(* IEC 61131-3 sources: SortJet_MasterSPS_Aufbau.fbsproj/10_Schnittstellen, 8 files *)

(* ---- Auftragswarteschlange_Fremdanlage_FB.fb.st ---- *)
(* METADATA
{
	"v3Meta": {
		"objectGuid": "565d8e9e-6f44-455e-86f5-d16ff6a06f95"
	}
}
*)
FUNCTION_BLOCK Auftragswarteschlange_Fremdanlage_FB
VAR_INPUT

  bpAktivieren     : BOOL := TRUE;
  bpWertAuslesen   : BOOL; // READ
  bpWerteSchreiben : BOOL; // WRITE
  bpReset          : BOOL; // RST

  // WORD
  ppEingabeWert : Schnittstelle_Auftragsdaten_ST;

END_VAR
VAR_OUTPUT
  // BOOLEAN
  bpWarteschlangeLeer  : BOOL := TRUE;
  bpWarteschlangeVoll  : BOOL;

  // STRUCT
  ppAusgabeWert  : Schnittstelle_Auftragsdaten_ST;

END_VAR
VAR

  // STRUCT
  awlWarteSchlange : ARRAY[0..cINDEX] OF Schnittstelle_Auftragsdaten_ST;

  // INT
  ilAktuellePosition  : INT; // pr
  ilLetztePosition    : INT; // pw

END_VAR

VAR CONSTANT
  cINDEX : INT := 5;    // WICHTIG: Aenderungen an diesem Wert aendert die Anzahl der Elemente in der Warteschlange [FIFO]
END_VAR
IF ( bpReset ) THEN
  ilLetztePosition := ilAktuellePosition := 0 ;
  bpWarteschlangeVoll := FALSE;
  bpWarteschlangeLeer := TRUE;

  bpReset := FALSE;

ELSIF ( bpAktivieren ) THEN

  IF (  NOT bpWarteschlangeLeer
       AND bpWertAuslesen )
  THEN
    ppAusgabeWert := awlWarteSchlange[ilAktuellePosition];
    ilAktuellePosition  := INCI(ilAktuellePosition,cINDEX);
    bpWarteschlangeLeer := ilAktuellePosition = ilLetztePosition;
    bpWarteschlangeVoll := FALSE;
    bpWertAuslesen      := FALSE;
  END_IF;

  IF (  NOT bpWarteschlangeVoll
       AND bpWerteSchreiben )
  THEN
    awlWarteSchlange[ilLetztePosition] := ppEingabeWert;
    ilLetztePosition    := INCI(ilLetztePosition,cINDEX);
    bpWarteschlangeVoll := ilLetztePosition = ilAktuellePosition;
    bpWarteschlangeLeer := FALSE;
    bpWerteSchreiben    := FALSE;
  END_IF;

END_IF;
END_FUNCTION_BLOCK

(* ---- Schnittstelle_Auslauf_ISO_FB.fb.st ---- *)
(* METADATA
{
	"v3Meta": {
		"objectGuid": "159241df-4e26-44a3-b242-7f4886765264"
	}
}
*)
FUNCTION_BLOCK Schnittstelle_Auslauf_ISO_FB EXTENDS Basic_Schnittstelle_FB_V01_00_00

VAR_INPUT
END_VAR
VAR_OUTPUT
END_VAR
VAR

  // STEPS
  steplStartIsolinie       : Steps_TE;

  // TRIGGER
  rtlAutomatik             : R_TRIG;
  rtlGlasAbruf             : R_TRIG;
  ftlGlasAbruf             : F_TRIG;

END_VAR

VAR_INPUT

  // HARDWARE EINGAENGE
  in_bGlasAbruf                 AT%I* : BOOL; // Signal von ISO-Linie
  in_bTransportRueckwaerts      AT%I* : BOOL; // Signal von ISO-Linie

  // ANALOGWERT
  in_wAnalogwertISOLinie        AT%I* : WORD; // Geschwindigkeit von der ISO-Linie

END_VAR

//-------------------------------------------------------------------------------------------------
// MASTER AUFRUFEN
//-------------------------------------------------------------------------------------------------
SUPER^(BasisStationsParameter := BasisStationsParameter);

//-------------------------------------------------------------------------------------------------
// BAUSTEIN: DEAKTIVIERUNG
//-------------------------------------------------------------------------------------------------
(* Hinweis:
   - Schnittstelle deaktiviert (MK bDeaktivieren): Baustein verlassen (Ausgaenge schaltet der Basis-Baustein ab)
*)
IF ( BasisStationsParameter.stMKs.bDeaktivieren ) THEN
  RETURN;
END_IF

//-------------------------------------------------------------------------------------------------
// BAUSTEIN: AKTIONEN
//-------------------------------------------------------------------------------------------------
CASE BasisStationsParameter.stMKs.stFremdanlage.eTypSchnittstelle OF

  //eGlaston:
  //  Glaston_Schnittstelle();

  eLISEC:
    Lisec_Schnittstelle();

  eFOREL:
    Forel_Schnittstelle();

  eHEGLA_SJ:
    Hegla_SJ_Schnittstelle();

END_CASE

// Meldung: Glas bereit, aber kein Abruf durch die Fremdanlage
Meldungen();

// Glaettung der Geschwindigkeit zur Sortierung
M_GeschwindigkeitGlaetten( rpMindestGeschwindigkeitsAenderung   := BasisStationsParameter.stMKs.stFremdanlage.rMindestGeschwindigkeitsAenderung,
                           tpMindestZeitZwischenGeschwAenderung := BasisStationsParameter.stMKs.stFremdanlage.tMindestZeitZwischenGeschwAenderung );

IF BasisStationsParameter.stMKs.stFremdanlage.bStationStatusZuGlasAbruf THEN
  Status_ISO_Linie();
END_IF

IF BasisStationsParameter.stMKs.stFremdanlage.bSignaleLoggen THEN
  Signal_Logger();
END_IF
END_FUNCTION_BLOCK

(* ---- Schnittstelle_Auslauf_Schneidanlage.fb.st ---- *)
(* METADATA
{
	"v3Meta": {
		"objectGuid": "5c116975-7ea8-4794-b20d-23cbba1de39f"
	}
}
*)
FUNCTION_BLOCK Schnittstelle_Auslauf_Schneidanlage EXTENDS Basic_Schnittstelle_FB_V01_00_00

VAR_INPUT
END_VAR

VAR_OUTPUT

  // Bool
  bpAnforderungSK : BOOL;
  bpGlasAbruf     : BOOL;

END_VAR

VAR

END_VAR

VAR_INPUT

  // HARDWARE EINGAENGE
  in_bGlasAbruf                 AT%I* : BOOL; // Signal von Schneidanlage
  in_bAnforderungSK             AT%I* : BOOL; // Signal von Schneidanlage

  out_bFreigabeSK               AT%Q* : BOOL; // Signal an Schneidanlage

END_VAR

//-------------------------------------------------------------------------------------------------
// MASTER AUFRUFEN
//-------------------------------------------------------------------------------------------------
SUPER^(BasisStationsParameter := BasisStationsParameter);

//-------------------------------------------------------------------------------------------------
// BAUSTEIN: DEAKTIVIERUNG
//-------------------------------------------------------------------------------------------------
(* Hinweis:
   - Schnittstelle deaktiviert (MK bDeaktivieren): Ausgaenge abschalten, Baustein verlassen
*)
IF ( BasisStationsParameter.stMKs.bDeaktivieren ) THEN
  out_bFreigabeSK := FALSE;
  bpAnforderungSK := FALSE;
  bpGlasAbruf     := FALSE;
  RETURN;
END_IF

//-------------------------------------------------------------------------------------------------
// BAUSTEIN: AKTIONEN
//-------------------------------------------------------------------------------------------------

Signalverarbeitung();
IF BasisStationsParameter.stMKs.stFremdanlage.bSignaleLoggen THEN
  Signal_Logger();
END_IF

//-------------------------------------------------------------------------------------------------
// STEUERUNG: HARDWARESCHNITTSTELLE
//-------------------------------------------------------------------------------------------------
blSenderGlasBereit := ( (*( BasisStationsParameter.bAutomatik )
                        AND*) NOT BasisStationsParameter.InGlasTransportVorgaenger[cWAND_1].bFehler )
                      AND ( BasisStationsParameter.InGlasTransportVorgaenger[cWAND_1].bBereitZumAustransport
                            OR BasisStationsParameter.bCheckMitVorgaenger[cWAND_1]
                            OR BasisStationsParameter.bCheckMitNachfolger[cWAND_1] );

bpAnforderungSK := in_bAnforderungSK OR bgVisu_Schnittstelle_Force_AnforderungSK[BasisStationsParameter.stMKs.stStationsNummern.NummerSPS];
bpGlasAbruf     := in_bGlasAbruf OR bgVisu_Schnittstelle_Force_GlasAbruf[BasisStationsParameter.stMKs.stStationsNummern.NummerSPS];

// SK-Freigabe an die Schneidanlage: nur auf Anforderung und bei Freigabe der Schnittstelle
out_bFreigabeSK := bpAnforderungSK AND BasisStationsParameter.stFreigabe.bAlles;

bgVisu_Schnittstelle_GlasAbruf[BasisStationsParameter.stMKs.stStationsNummern.NummerSPS]     := in_bGlasAbruf OR bgVisu_Schnittstelle_Force_GlasAbruf[BasisStationsParameter.stMKs.stStationsNummern.NummerSPS];
bgVisu_Schnittstelle_AnforderungSK[BasisStationsParameter.stMKs.stStationsNummern.NummerSPS] := in_bAnforderungSK OR bgVisu_Schnittstelle_Force_AnforderungSK[BasisStationsParameter.stMKs.stStationsNummern.NummerSPS];
bgVisu_Schnittstelle_FreigabeSK[BasisStationsParameter.stMKs.stStationsNummern.NummerSPS]    := out_bFreigabeSK;
END_FUNCTION_BLOCK

(* ---- Schnittstelle_Auslauflinie_Glaston_Koppler_FB.fb.st ---- *)
(* METADATA
{
	"v3Meta": {
		"objectGuid": "1b8cd41b-c6ec-4747-8cfe-b17b04789a14"
	}
}
*)
FUNCTION_BLOCK Schnittstelle_Auslauflinie_Glaston_Koppler_FB  EXTENDS Basic_Schnittstelle_FB_V01_00_00

VAR_INPUT

  // BOOL
  bpAuftragsdatenVorhanden  : BOOL;

  // STRUCT
  Auftragsdaten             : Schnittstelle_Auftragsdaten_ST;

END_VAR
VAR_OUTPUT

END_VAR
VAR

  // BOOL
  bpDatenformatASCII                      : BOOL := TRUE;
  blLiveCounterGueltig                    : BOOL;
  blFehlermeldungGenerierenKommunikation  : BOOL;
  blFehlermeldungGenerierenAuftragsdaten  : BOOL;
  bpFehlerMeldungDeaktiviert              : BOOL := FALSE;

  // BYTE
  aOutByteLadeID             : ARRAY [0..15] OF BYTE; // Visualisierung: Lade-ID byteweise

  // WORD
  wlVerbindungsVersuche      : WORD;
  wlLiveCounterSortJet       : WORD;
  wlLiveCounterFremdanlage   : WORD;
  wlTempEmpfaengerSignale    : WORD;
  wlTempSenderSignale        : WORD;
  wlOutSignale               : WORD;
  wlInSignale                : WORD;

  // DWORD
  dwlGeschwindigkeit         : DWORD;                   // Geschwindigkeit des Empfaengers [mm/s], ggf. geswappt
  adwlLadeID                 : ARRAY [0..3] OF DWORD;   // Lade-ID (= Scheiben-ID 1), ggf. geswappt

  // INT
  ilIndex                    : INT;

  // TRIGGER
  ftlGlasBereit                           : F_TRIG; // Hinweis: Glas-Sender besitzt noch einen aktiven Transport-Zustand
  ftlFremdanlageDatenVerarbeitet          : F_TRIG;
  rtlFehlermeldungGenerierenAuftragsdaten : R_TRIG;
  rtlFehlermeldungGenerierenKommunikation : R_TRIG;

  // TIMER
  tonlZeitLiveCounterNichtAequivalent     : TON;
  tonlZeitLiveCounterInkrementieren       : TON;
  tonlZeitAuftragsdatenNichtAequivalent   : TON;
  tonlManuellerModus                      : TON;
  tonlAuftragdatenVorhanden               : TON;

  // STRING
  strScheibenID  : STRING;

  // STRUCT
  stlAuftragsdatenLeer : Schnittstelle_Auftragsdaten_ST; // Leere Auftragsdaten zum Loeschen beim Reset

  // REFERENZ
  stlVorgaenger  : REFERENCE TO StationBasisParameter_ST; // SortJet- Station vor der Schnittstelle (SF/SB)

END_VAR

VAR

  // STEPS
  steplStartIsolinie                                     : Steps_TE;

  // TRIGGER
  rtlAutomatik                                           : R_TRIG;
  rtlGlasAbruf                                           : R_TRIG;
  ftlGlasAbruf                                           : F_TRIG;

  // HARDWARE EINGAENGE KOPPLER (Hegla Schnittstellenbeschreibung V4.0, Empfaenger -> Sender)
  in_wEmpfaengerLiveCounter                     AT %I*   : WORD;                  // Wort 0     LC: gespiegelter LiveCounter
  in_awEmpfaengerLadeIDGespiegelt               AT %I*   : ARRAY [1..8] OF WORD;  // Wort 1..8  ID: gespiegelte Lade-ID
  in_wEmpfaengerSignale                         AT %I*   : WORD;                  // Wort 49    Signale
  in_dwEmpfaengerGeschwindigkeit                AT %I*   : DWORD;                 // Wort 50    GE: Geschwindigkeit [mm/s]
  in_wEmpfaengerRampe                           AT %I*   : WORD;                  // Wort 52    RA [Option]: Rampe [mm/s²], nur Anzeige

  in_bEmpfaengerAuftragsdatenErhalten                    : BOOL; // 49.0 AG
  in_bEmpfaengerBereitZumEintransport                    : BOOL; // 49.1 GA
  in_bEmpfaengerNothalt                                  : BOOL; // 49.3 NA  [Option] nur Anzeige
  in_bEmpfaengerAnforderungDurchgangOeffnen              : BOOL; // 49.4 ADO [Option] nur Anzeige
  in_bEmpfaengerQuittungDurchgangOeffnen                 : BOOL; // 49.5 ADQ [Option] nur Anzeige
  in_bEmpfaengerStationFrei                              : BOOL; // 49.6 SF  [Option]
  in_bEmpfaengerStationBeladen                           : BOOL; // 49.7 SB  [Option]
  in_bEmpfaengerUebernahmeposition                       : BOOL; // 49.8 UP  [Option] nur Anzeige

  // HARDWARE AUSGAENGE KOPPLER (Hegla Schnittstellenbeschreibung V4.0, Sender -> Empfaenger)
  out_wSenderLiveCounter                     AT %Q*      : WORD;                  // Wort 0     LC: LiveCounter
  out_awSenderLadeID                         AT %Q*      : ARRAY [1..8] OF WORD;  // Wort 1..8  ID: Lade-ID (16 ASCII- Zeichen)
  out_wSenderSignale                         AT %Q*      : WORD;                  // Wort 50    Signale

  out_bSenderAuftragdatenVorhanden                       : BOOL; // 50.0 AV
  out_bSenderAuftragdatenPlausibel                       : BOOL; // 50.1 AP
  out_bSenderManuelleBeladung                            : BOOL; // 50.2 HB [Option] SortJet sendet immer mit Lade-ID
  out_bSensorAuslauf                                     : BOOL; // 50.6 SA [Option]
  out_bSenderStationFrei                                 : BOOL; // 50.7 SF [Option] Vorgaengerstation frei
  out_bSenderStationBeladen                              : BOOL; // 50.8 SB [Option] Vorgaengerstation belegt
  out_bSenderForm                                        : BOOL; // 50.9 FG [Option] Scheibe ist ein Modell

END_VAR
VAR CONSTANT

  // WORD
  cVERBINDUNGSVERSUCHE_BIS_FEHLER  : WORD := 5;         // WICHTIG: Aenderung an diesem Wert veraendert das Verhalten ab wieviel Kommunikations-Versuchen wann ein Fehler ausgegeben wird

  // INT
  cWERTEBREICH_INT                 : INT  := 32767; // WICHTIG: Aenderung an diesem Wert aendert den Wertebereich eines INTs [positiver Wertebereich]
  cWERTEBREICH_WORD                : WORD := 32767; // WICHTIG: Aenderung an diesem Wert aendert den Wertebereich eines INTs [positiver Wertebereich]

  // TIME
  cZEIT_AUFTRAGSDATEN_GUELTIG                : TIME :=T#5s;         // WICHTIG: Aenderung an diesem Wert aendert die Zeit ab wann ein Fehlergeneriert wird [s]
  cZEIT_GESPIEGELTE_AUFTRAGSDATEN_UNGUELTIG  : TIME :=T#5s;         // WICHTIG: Aenderung an diesem Wert aendert die Zeit ab wann ein Fehlergeneriert wird [s]
  cZEIT_MANUELLER_MODUS_SIGNAL               : TIME :=T#10s;
  cZEIT_LIVECOUNTER_INKREMENTIEREN           : TIME :=T#250ms;
  cZEIT_LIVECOUNTER_NICHT_GUELTIG            : TIME :=T#1500ms;

END_VAR
//-------------------------------------------------------------------------------------------------
// MASTER AUFRUFEN
//-------------------------------------------------------------------------------------------------
SUPER^(BasisStationsParameter := BasisStationsParameter);

//-------------------------------------------------------------------------------------------------
// BAUSTEIN: INITIALISIERUNG
//-------------------------------------------------------------------------------------------------
IF ( blErsterZyklus  ) THEN
  blErsterZyklus := FALSE;

  bpAuftragsdatenVorhanden      := FALSE;
  AuftragsSpeicher.bpAktivieren := TRUE;

END_IF

//-------------------------------------------------------------------------------------------------
// BAUSTEIN: DEAKTIVIERUNG
//-------------------------------------------------------------------------------------------------
(* Hinweis:
   - Schnittstelle deaktiviert (MK bDeaktivieren): Signalwort zum Empfaenger nullen, Baustein verlassen
     (der LiveCounter bleibt stehen -> Empfaenger erkennt die fehlende Kommunikation)
*)
IF ( BasisStationsParameter.stMKs.bDeaktivieren ) THEN
  out_wSenderSignale := 0;
  RETURN;
END_IF

//-------------------------------------------------------------------------------------------------
// TIMER
//-------------------------------------------------------------------------------------------------
(* Hinweis:
   - Zeitlicheueberwachung der Kommunikation
*)
tonlZeitLiveCounterNichtAequivalent( IN := NOT blLiveCounterGueltig,
                                     PT := cZEIT_LIVECOUNTER_NICHT_GUELTIG );

//-------------------------------------------------------------------------------------------------
// AKTIONEN
//-------------------------------------------------------------------------------------------------
LiveCounter();
Meldungen();
AuftragsdatenVerwaltung();
Auswertung();
Signalverarbeitung();
M_GeschwindigkeitGlaetten( rpMindestGeschwindigkeitsAenderung   := BasisStationsParameter.stMKs.stFremdanlage.rMindestGeschwindigkeitsAenderung,
                           tpMindestZeitZwischenGeschwAenderung := BasisStationsParameter.stMKs.stFremdanlage.tMindestZeitZwischenGeschwAenderung );
Status_ISO_Linie();

IF BasisStationsParameter.stMKs.stFremdanlage.bSignaleLoggen THEN
  Signal_Logger();
END_IF

//-------------------------------------------------------------------------------------------------
// RESET
//-------------------------------------------------------------------------------------------------
// Fehlverhalten:
//   - Anstehenden Fehler zuruecksetzen
IF ( BasisStationsParameter.bReset ) THEN

  out_bSenderAuftragdatenPlausibel := FALSE;
  out_bSenderAuftragdatenVorhanden := FALSE;

  bpAuftragsdatenVorhanden               := FALSE;
  blFehlermeldungGenerierenKommunikation := FALSE;
  blFehlermeldungGenerierenAuftragsdaten := FALSE;

  BasisStationsParameter.bReset := FALSE;

  // Auftragsdaten komplett loeschen
  Auftragsdaten := stlAuftragsdatenLeer;

END_IF

//-------------------------------------------------------------------------------------------------
// Aufrufe
//-------------------------------------------------------------------------------------------------
Horn( bpAktiv := bgHornAktivieren );
END_FUNCTION_BLOCK

(* ---- Schnittstelle_Einlauf_HeglaBrechanlage_FB.fb.st ---- *)
(* METADATA
{
	"v3Meta": {
		"objectGuid": "887b7e5f-63a1-4543-befe-d3acd4ce4d49"
	}
}
*)
{attribute 'excludefrombuild'}
FUNCTION_BLOCK Schnittstelle_Einlauf_HeglaBrechanlage_FB
(*
//=================================================================================================
// !!! TODO !!! TODO !!! TODO !!! TODO !!! TODO !!! TODO !!! TODO !!! TODO !!! TODO !!! TODO !!!
//=================================================================================================
// - Dieser Baustein erbt NICHT von Basic_Schnittstelle_FB_V01_00_00.
// - Er ist nicht instanziiert und nicht im Build (excludefrombuild).
// - Vor der Verwendung auf die Basis-Schnittstelle umstellen:
//     EXTENDS, SUPER^, Reset und Meldungen der Basis nutzen, danach testen.
//=================================================================================================
*)
VAR_INPUT

  // BOOL
  bpStarteReset                 : BOOL;
  bpAnforderungSK               : BOOL;

  // STRUCT
  InGlasTransportNachfolger     : Interface_GlasTransport;
  stStationsNummern             : Station_ST;

  // POINTER
  ppParameterBaustein : REFERENCE TO Parameter_Schnittstelle;

END_VAR
VAR_OUTPUT

  // STRUCT
  OutGlasTransport : Interface_GlasTransport; // STRUKTUR: Informationen ueber den Aus- Ein- Transport WAND 1

END_VAR
VAR

  // BOOL
  blErsterZyklus          : BOOL := TRUE;

  // TIMER
  tonlMeldungGenerierenGLassenderNichtBereit : TON;// EINSCHALTVERZOEGERUNG

END_VAR
VAR

  // HARDWARE EINGAENGE
  in_bGlasBereit                AT %I* : BOOL; // Glas auf Brechanlage bereit zum Austransport
  in_bFreigabeSK                AT %I* : BOOL; // Freigabe zum SK 2 öffnen
  in_bAnlageEingeschaltet       AT %I* : BOOL; // Signal zum Zustand der Brechanlage, ob Eingeschaltet oder nicht
  in_bSensorAuslauf             AT %I* : BOOL; // Auslaufsensor (letzter Sensor vor Übergabe) der Brechanlage
  in_bBypassMode                AT %I* : BOOL; // ByPass an Brechanlage aktiv: Übergroße Scheiben für die Brechanlage müssen ohne Analogwert gefahren werden ; Festgesetzte Geschw. 20m/min zwischen Brechanlage und SortJet

  // HARDWARE AUSGAENGE
  out_bGlasAbruf                AT %Q* : BOOL; // Glas Abruf zur Brechanlage, sofern Glas Bereit ist
  out_bAnforderungSK            AT %Q* : BOOL; // Anforderung zum öffnen des 2. SK - Brechanlage muss in sichere Stop-Position fahren und freigeben
  out_bSensorEinlauf            AT %Q* : BOOL; // Erster Sensor am RKT
  out_bReserve                  AT %Q* : BOOL; // Optional

  out_wSpeed                    AT %Q* : WORD;

END_VAR
IF ( blErsterZyklus ) THEN
  blErsterZyklus:=FALSE;

  (* Wichtig:
     - Pointer Initialisieren [Null-Pointer-Exception]
  *)
  InGlasTransportNachfolger  := NullReferenzGlasTransport;
  OutGlasTransport           := NullReferenzGlasTransport;

  (* Hinweis:
     - Basis- Pointer uebergeben
  *)
  ppParameterBaustein  := ADR( apgMKSchnittstelle_Einlauflinie[stStationsNummern.NummerSPS]);

END_IF

//-------------------------------------------------------------------------------------------------
// BAUSTEIN: SCHNITTSTELLE
//-------------------------------------------------------------------------------------------------
(* Hinweis:
   - Abhandlung des Ein-Aus- Transports [Setzen der Variablen das man bereit ist zum Glastransport]
*)
OutGlasTransport.stStationsNummern      := stStationsNummern;
OutGlasTransport.wStationsTyp           := eFremdanlage;
OutGlasTransport.bEinlaufsensor         := ADR(bgFALSE);
OutGlasTransport.bAuslaufsensor         := ADR(in_bSensorAuslauf);
OutGlasTransport.bBereitZumAustransport := ADR(in_bGlasBereit);
OutGlasTransport.bBereitZumEintransport := ADR(bgFALSE);
OutGlasTransport.bFehler                := ADR(bgFALSE);
OutGlasTransport.rGeschwindigkeit       := ADR(rgNull);

//-------------------------------------------------------------------------------------------------
// BAUSTEIN: AKTIONEN
//-------------------------------------------------------------------------------------------------

CASE ppParameterBaustein.eTypSchnittstelle OF

  eHEGLA_BREAK:
    HeglaBrechanlage_Schnittstelle();

END_CASE

// Aktion:
//   - Reset
Reset();

//-------------------------------------------------------------------------------------------------
// BAUSTEIN: MELDUNGEN
//-------------------------------------------------------------------------------------------------

(* Hinweis:
   - Meldungs Sender nicht bereit
*)
tonlMeldungGenerierenGLassenderNichtBereit( IN :=  InGlasTransportNachfolger.AND NOT in_bGlasBereit,
                                            PT :=  t#30s );

WatchIo( tonlMeldungGenerierenGLassenderNichtBereit.Q , ( ppParameterBaustein.wMeldungsNummer ) );
END_FUNCTION_BLOCK

(* ---- Schnittstelle_Einlauf_Portale.fb.st ---- *)
(* METADATA
{
	"v3Meta": {
		"objectGuid": "1983d120-77fe-4da5-a5d1-bf513123edf7"
	}
}
*)
FUNCTION_BLOCK Schnittstelle_Einlauf_Portale EXTENDS Basic_Schnittstelle_FB_V01_00_00
VAR_INPUT

  // HARDWARE EINGAENGE
  in_bGlasAufgestellt                     AT %I* : BOOL;

END_VAR

VAR_OUTPUT

  // HARDWARE AUSGAENGE
  out_bBereitZumAufstellen               AT %Q* : BOOL;

END_VAR

// Schnittstelle zu den Portalen (Glas aufstellen)
// - "out_bBereitZumAufstellen": die Folgestation ist bereit zum Eintransport, das Portal darf Glas aufstellen
// - "in_bGlasAufgestellt": das Portal hat Glas aufgestellt, die Folgestation startet den Eintransport

//-------------------------------------------------------------------------------------------------
// MASTER AUFRUFEN
//-------------------------------------------------------------------------------------------------
SUPER^(BasisStationsParameter := BasisStationsParameter);

//-------------------------------------------------------------------------------------------------
// BAUSTEIN: DEAKTIVIERUNG
//-------------------------------------------------------------------------------------------------
(* Hinweis:
   - Schnittstelle deaktiviert (MK bDeaktivieren): Ausgaenge abschalten, Baustein verlassen
*)
IF ( BasisStationsParameter.stMKs.bDeaktivieren ) THEN
  out_bBereitZumAufstellen := FALSE;
  RETURN;
END_IF

IF BasisStationsParameter.stMKs.stFremdanlage.bSignaleLoggen THEN
  Signal_Logger();
END_IF

//-------------------------------------------------------------------------------------------------
// SCHNITTSTELLE
//-------------------------------------------------------------------------------------------------
// Signale vom Portal
blBereitZumAustransport := in_bGlasAufgestellt OR bgVisu_Schnittstelle_Einlauf_Force_GlasBereit[BasisStationsParameter.stMKs.stStationsNummern.NummerSPS];

//-------------------------------------------------------------------------------------------------
// MELDUNGEN
//-------------------------------------------------------------------------------------------------
// Portal hat Glas aufgestellt, die Station ist aber 30 s nicht bereit zum Eintransport [wMeldungsNummer + 2]
WatchIoControl( T#30S,
                BasisStationsParameter.stMKs.wMeldungsNummer + 2,
                blBereitZumAustransport AND NOT BasisStationsParameter.InGlasTransportNachfolger[cWAND_1].bBereitZumEintransport );

//-------------------------------------------------------------------------------------------------
// AUSGAENGE
//-------------------------------------------------------------------------------------------------
// Signale zum Portal
out_bBereitZumAufstellen := BasisStationsParameter.InGlasTransportNachfolger[cWAND_1].bBereitZumEintransport;

//-------------------------------------------------------------------------------------------------
// VISU
//-------------------------------------------------------------------------------------------------
bgVisu_Schnittstelle_Einlauf_Status_GlasBereit[BasisStationsParameter.stMKs.stStationsNummern.NummerSPS]   := BasisStationsParameter.OutGlasTransport[cWAND_1].bBereitZumAustransport;
bgVisu_Schnittstelle_Status_BereitZumEintrasport[BasisStationsParameter.stMKs.stStationsNummern.NummerSPS] := out_bBereitZumAufstellen;
END_FUNCTION_BLOCK

(* ---- Schnittstelle_Einlauf_VSG.fb.st ---- *)
(* METADATA
{
	"v3Meta": {
		"objectGuid": "fbbba330-556c-41e3-bb2c-ea5fa1aaa6e1"
	}
}
*)
FUNCTION_BLOCK Schnittstelle_Einlauf_VSG EXTENDS Basic_Schnittstelle_FB_V01_00_00
VAR_INPUT

END_VAR
VAR_OUTPUT

  // STRUCT
  OutGlasTransport   : Interface_LTR_VSG; // Signale zum LTR

END_VAR

VAR_INPUT

  // HARDWARE EINGAENGE
  in_bGlasBereit                          AT %I* : BOOL;
  in_bAutomatikBetrieb                    AT %I* : BOOL; // Scheiben werden automatisch eintransportiert

END_VAR

VAR_OUTPUT
  // HARDWARE AUSGAENGE
  out_bEinlaufsensor                      AT %Q* : BOOL;
  out_bBereitZumEintrasport               AT %Q* : BOOL;

END_VAR

// Schnittstelle zwischen LTR und VSG Anlage
// Sobald wir einen Anlageauftrag bekommen und das Signal "in_bAutomatikBetrieb" ansteht, gehen wir in Eintrasport.
// Dort setzen wir "out_bBereitZumEintrasport" und warten bis das Signal "in_bGlasBereit" ansteht. Dieses wird von
// der VSG gesetzt wenn Glas bereit liegt und die Riemen in SlaveMode sind. Wir starten dann denn Eintransport.
// Der SlaveMode bleibt so lange aktiv, bis wir das Signal "out_bBereitZumEintrasport" wegnehmen.

//-------------------------------------------------------------------------------------------------
// MASTER AUFRUFEN
//-------------------------------------------------------------------------------------------------
SUPER^(BasisStationsParameter := BasisStationsParameter);

//-------------------------------------------------------------------------------------------------
// BAUSTEIN: DEAKTIVIERUNG
//-------------------------------------------------------------------------------------------------
(* Hinweis:
   - Schnittstelle deaktiviert (MK bDeaktivieren): Ausgaenge abschalten, Baustein verlassen
*)
IF ( BasisStationsParameter.stMKs.bDeaktivieren ) THEN
  out_bEinlaufsensor        := FALSE;
  out_bBereitZumEintrasport := FALSE;
  RETURN;
END_IF

IF BasisStationsParameter.stMKs.stFremdanlage.bSignaleLoggen THEN
  Signal_Logger();
END_IF

//-------------------------------------------------------------------------------------------------
// SCHNITTSTELLE
//-------------------------------------------------------------------------------------------------
// Signale von der VSG
blBereitZumAustransport := in_bGlasBereit OR bgVisu_Schnittstelle_Einlauf_Force_GlasBereit[BasisStationsParameter.stMKs.stStationsNummern.NummerSPS];
blAutomatikBetriebAktiv := in_bAutomatikBetrieb OR bgVisu_Schnittstelle_Force_AutomatikBetrieb[BasisStationsParameter.stMKs.stStationsNummern.NummerSPS];;

//-------------------------------------------------------------------------------------------------
// MELDUNGEN
//-------------------------------------------------------------------------------------------------
// VSG-Linie hat Glas bereit, die Station ist aber 30 s nicht bereit zum Eintransport [wMeldungsNummer + 2]
WatchIoControl( T#30S,
                BasisStationsParameter.stMKs.wMeldungsNummer + 2,
                blBereitZumAustransport AND NOT BasisStationsParameter.InGlasTransportNachfolger[cWAND_1].bBereitZumEintransport );

//-------------------------------------------------------------------------------------------------
// AUSGAENGE
//-------------------------------------------------------------------------------------------------
// Signale zur VSG
out_bEinlaufsensor        := BasisStationsParameter.InGlasTransportNachfolger[cWAND_1].bEinlaufsensor;
out_bBereitZumEintrasport := BasisStationsParameter.InGlasTransportNachfolger[cWAND_1].bBereitZumEintransport;

//-------------------------------------------------------------------------------------------------
// VISU
//-------------------------------------------------------------------------------------------------
bgVisu_Schnittstelle_Einlauf_Status_GlasBereit[BasisStationsParameter.stMKs.stStationsNummern.NummerSPS]   := BasisStationsParameter.OutGlasTransport[cWAND_1].bBereitZumAustransport;
bgVisu_Schnittstelle_Status_AutomatikBetrieb[BasisStationsParameter.stMKs.stStationsNummern.NummerSPS]     := BasisStationsParameter.OutGlasTransport[cWAND_1].bAutomatikBetriebAktiv;
bgVisu_Schnittstelle_Status_Einlaufsensor[BasisStationsParameter.stMKs.stStationsNummern.NummerSPS]        := out_bEinlaufsensor;
bgVisu_Schnittstelle_Status_BereitZumEintrasport[BasisStationsParameter.stMKs.stStationsNummern.NummerSPS] := out_bBereitZumEintrasport;
END_FUNCTION_BLOCK

(* ---- Schnittstelle_Einlauflinie_FB.fb.st ---- *)
(* METADATA
{
	"v3Meta": {
		"objectGuid": "583875e0-db52-49ee-af9c-0f6353b622c9"
	}
}
*)
{attribute 'excludefrombuild'}
FUNCTION_BLOCK Schnittstelle_Einlauflinie_FB
(*
//=================================================================================================
// !!! TODO !!! TODO !!! TODO !!! TODO !!! TODO !!! TODO !!! TODO !!! TODO !!! TODO !!! TODO !!!
//=================================================================================================
// - Dieser Baustein ist UNFERTIG.
// - Er erbt NICHT von Basic_Schnittstelle_FB_V01_00_00.
// - Er ist nicht instanziiert und nicht im Build (excludefrombuild).
// - Vor der Verwendung fertigstellen und auf die Basis-Schnittstelle umstellen:
//     EXTENDS, SUPER^, Reset und Meldungen der Basis nutzen, danach testen.
//=================================================================================================
*)
VAR_INPUT

  // BOOLEAN
  bpReset                         : BOOL;
  bpAktivieren                    : BOOL := TRUE;
  bpSortierungInAutomatik         : BOOL; // [STATUS] Status der Sortierung -> Automatikbetrieb
  bpNotHaltAusgeloest              : BOOL := FALSE;
  bpDatenformatASCII              : BOOL := TRUE;

  // STRUCT
  InGlasTransport    : Interface_GlasTransport;        // STRUKTUR: Informationen ueber den Aus- Ein- Transport WAND 1
  Auftragsdaten      : Schnittstelle_Auftragsdaten_ST; // STRUKTUR: Auftragsdaten fuer die Fremdanlage [ScheibenID , Auftragsnummer , etc. ]
  stStationsNummern  : Station_ST;

  // POINTER
  ppParameterBaustein : REFERENCE TO Parameter_Schnittstelle;

END_VAR
VAR_OUTPUT

  // BOOLEAN
  bpFehler      : BOOL;

  // STRUCT
  OutGlasTransport   : Interface_GlasTransport; // STRUKTUR: Informationen ueber den Aus- Ein- Transport WAND 1

END_VAR
VAR

  // BOOLEAN
  blErsterZyklus                          : BOOL := TRUE;  // Initialisierung
  blAuftragAktiv                          : BOOL := FALSE;
  blFehlermeldungGenerierenKommunikation  : BOOL;
  blFremdanlageBereitZumTransport         : BOOL := FALSE;
  blAuftragsdatenNachrichtGenerieren      : BOOL;

  // BYTE
  aInByteAuftragsdatenScheibenID_1_0     : ARRAY [0..3] OF BYTE;
  aInByteAuftragsdatenScheibenID_1_1     : ARRAY [0..3] OF BYTE;
  aInByteAuftragsdatenScheibenID_1_2     : ARRAY [0..3] OF BYTE;
  aInByteAuftragsdatenScheibenID_1_3     : ARRAY [0..3] OF BYTE;
  aInByteSwapAuftragsdatenScheibenID_1_0 : ARRAY [0..3] OF BYTE;
  aInByteSwapAuftragsdatenScheibenID_1_1 : ARRAY [0..3] OF BYTE;
  aInByteSwapAuftragsdatenScheibenID_1_2 : ARRAY [0..3] OF BYTE;
  aInByteSwapAuftragsdatenScheibenID_1_3 : ARRAY [0..3] OF BYTE;

  // WORD
  wlMerkerLiveCounterSender             : WORD;
  wlLiveCounterSender                   : WORD;

  // INT
  ilIndex  : INT;

  // DWORD
  aInDWordAuftragsdatenScheibenID : ARRAY [0..3] OF DWORD;

  // STRING
  strScheibenID : STRING;

  // TRIGGER
  rtlAutomatikActiv                       : R_TRIG;
  rtlFehlermeldungGenerierenKommunikation : R_TRIG;
  rtlAuftragsdatenPlausibel               : R_TRIG;
  ftlAuftragsdatenVorhanden               : F_TRIG;

  // TIMER
  tonlUeberwachungLiveCounter            : TON; // EINSCHALTVERZOEGERUNG

END_VAR
VAR

  // HARDWARE EINGAENGE
  in_stSenderAuftragsdaten                      AT %I* : Schnittstelle_ScheibenIDs;  // HINWEIS: PROFIBUS- Schnittstelle
  in_wSenderLiveCounter                         AT %I* : WORD;
  in_bSenderAuftragdatenVorhanden               AT %I* : BOOL; // HINWEIS: PROFIBUS- Schnittstelle
  in_bsenderAuftragdatenPlausibel               AT %I* : BOOL; // HINWEIS: PROFIBUS- Schnittstelle
  in_bSenderBereit                              AT %I* : BOOL; // HINWEIS: PROFIBUS- Schnittstelle
  in_bSenderGlasBereit                          AT %I* : BOOL; // HINWEIS: PROFIBUS- Schnittstelle -> Glas bereit zum Eintransport [Sortierung zur Fremdanlage]
  in_bSenderSensorAuslauf                       AT %I* : BOOL; // HINWEIS: SPS- Eingang des Sensors auf die PROFIBUS- Schnittstelle schreiben [Sortierung zur Fremdanlage]
  in_bSenderScheibeManuellAnlegen               AT %I* : BOOL; // HINWEIS: PROFIBUS- Schnittstelle
  in_wSenderAnzahlScheiben                      AT %I* : WORD := 0;

  // HARDWARE AUSGAENGE
  out_wEmpfaengerLiveCounter                    AT %Q* : WORD; // HINWEIS: ANYBUS - Schnittstelle
  out_stEmpfaengerAuftragsdatenGespiegelt       AT %Q* : Schnittstelle_ScheibenIDs; // HINWEIS: PROFIBUS- Schnittstelle
  out_bEmpfaengerAuftragsdatenErhalten          AT %Q* : BOOL; // HINWEIS: PROFIBUS- Schnittstelle
  out_bEmpfaengerGlasAbruf                      AT %Q* : BOOL;
  out_bEmpfaengerSensorEinlauf                  AT %Q* : BOOL;
  out_bEmpfaengerNotHaltAusgeloest               AT %Q* : BOOL;
  out_rEmpfaengerGeschwindigkeit                AT %Q* : REAL := REAL#0;
  out_bEmpfaengerBetriebsbereit                        : BOOL;
  out_bEmpfaengerGlasuebernommen                       : BOOL;

END_VAR
VAR CONSTANT

  // TIME
  cZEIT_UEBERWACHUNG_LIVECOUNTER    : TIME :=T#5s; // WICHTIG: Aenderung an diesem Wert aendert die Zeit ab wann ein Fehlergeneriert wird [s]

END_VAR
(* Hinweis:
   - Dieser Baustein bildet das Interface zu einer Fremdanlage
     => Verarbeitung der Signale [ Bereit zum Eintransport | Bereit zum Austransport ]
*)

//-------------------------------------------------------------------------------------------------
// BAUSTEIN: INITIALISIERUNG
//-------------------------------------------------------------------------------------------------
IF ( blErsterZyklus  ) THEN
  blErsterZyklus := FALSE;

  (* Hinweis [OPTIONAL]:
     - Auftragsdaten nullen
  *)
  out_stEmpfaengerAuftragsdatenGespiegelt := NullReferenzAuftragsdatenFremdanlage.stScheibenID;

  (* Wichtig:
     - Pointer Initialisieren [Null-Pointer-Exception]
  *)
  InGlasTransport := NullReferenzGlasTransport;

  (* Hinweis:
     - Basis- Pointer uebergeben
  *)
  ppParameterBaustein  := ADR( apgMKSchnittstelle_Einlauflinie[stStationsNummern.NummerSPS]);

END_IF

//-------------------------------------------------------------------------------------------------
// SCHNITTSTELLE
//-------------------------------------------------------------------------------------------------
(* Hinweis:
   - Abhandlung des Ein-Aus- Transports [Setzen der Variablen das man bereit ist zum Glastransport]
*)
OutGlasTransport.stStationsNummern      := stStationsNummern;
OutGlasTransport.wStationsTyp           := eFremdanlage;
OutGlasTransport.bEinlaufsensor         := ADR( bgFalse );
OutGlasTransport.bAuslaufsensor         := ADR( in_bSenderSensorAuslauf );
OutGlasTransport.bBereitZumAustransport := ADR( blFremdanlageBereitZumTransport );
OutGlasTransport.bBereitZumEintransport := ADR( blFremdanlageBereitZumTransport );
OutGlasTransport.rGeschwindigkeit       := ADR( rgMkAutoGeschwindigkeitFremdanlage );
OutGlasTransport.bFehler                := ADR( bpFehler );

//-------------------------------------------------------------------------------------------------
// Deaktivierung
//-------------------------------------------------------------------------------------------------
IF ( NOT bpAktivieren ) THEN
  RETURN;
END_IF

//-------------------------------------------------------------------------------------------------
// SIGNALVERARBEITUNG [HARDWARE EIN- AUS- GAENGE | ETC. ]
//-------------------------------------------------------------------------------------------------
(* Hinweis:
   - Signal das der Sender bereit fuer den Transport ist
*)
blFremdanlageBereitZumTransport := (     in_bSenderBereit
                                     AND in_bSenderGlasBereit );

(* Hinweis:
   - Glas Abrufen von der Fremdanlage
*)
out_bEmpfaengerGlasAbruf := (         InGlasTransport.bBereitZumEintransport^
                              AND NOT bgVisu_Schnittstelle_Force_EmpfaengerFreiInGlasTransport.bFehler^ );

(* Hinweis:
   - Geschwindigkeit
*)
out_rEmpfaengerGeschwindigkeit := InGlasTransport.rGeschwindigkeit;

(* Hinweis:
   - Der Auslaufsensor der Vorgaengerstation uebergeben
*)
out_bEmpfaengerSensorEinlauf := InGlasTransport.bEinlaufsensor;

(* Hinweis:
   - NotAus
*)
out_bEmpfaengerNotHaltAusgeloest := bpNotHaltAusgeloest;

//-------------------------------------------------------------------------------------------------
// AKTIONEN
//-------------------------------------------------------------------------------------------------
(* Hinweis:
   - Baustein-Aktionen
*)
LiveCounter();
Ausnahmesituation();
AuftragsdatenVerwaltung();
Auswertung();

//-------------------------------------------------------------------------------------------------
// RESET
//-------------------------------------------------------------------------------------------------
// Fehlverhalten:
//   - Anstehenden Fehler zuruecksetzen
IF ( bpReset ) THEN

  bpFehler       := FALSE;
  blAuftragAktiv := FALSE;

  blFehlermeldungGenerierenKommunikation := FALSE;

  bpReset := FALSE;

END_IF
END_FUNCTION_BLOCK
